FUNCTION_BLOCK TestingSequence (* Basic Function Block Type *)
  (* Standard: 61499-2 *)
  (* Version 0.0, 11/16/2026, Sandeep Patil, Flexbridge AB, Template *)
  PACKAGE Flexbridge.FestoMPS400;
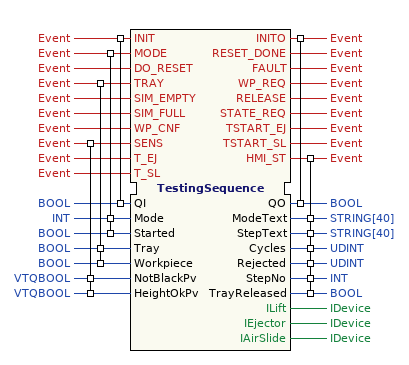
  EVENT_INPUT
    INIT WITH QI; (* Initialisation request *)
    MODE WITH Mode, Started; (* Station mode changed (StationMode) *)
    DO_RESET; (* Run the reset sequence (StationMode) *)
    TRAY WITH Tray, Workpiece; (* Tray state at interface 1 (conveyor waypoint, IWaypoint) *)
    SIM_EMPTY; (* Stand-in: an empty tray has arrived (HMI button) *)
    SIM_FULL; (* Stand-in: a tray with a workpiece has arrived (HMI button) *)
    WP_CNF; (* Distributing has handed a workpiece over (IWorkpieceSupply) *)
    SENS WITH NotBlackPv, HeightOkPv; (* Colour or height sensor changed *)
    T_EJ; (* Ejector time over (EjectTimer) *)
    T_SL; (* Air slide time over (SlideTimer) *)
  END_EVENT
  EVENT_OUTPUT
    INITO WITH QO; (* Initialisation confirm *)
    RESET_DONE; (* Reset sequence finished (StationMode) *)
    FAULT; (* Stopped on a device fault (StationMode) *)
    WP_REQ; (* Ask Distributing for a workpiece (IWorkpieceSupply) *)
    RELEASE; (* Release the tray (IWaypoint) *)
    STATE_REQ; (* Ask the waypoint for the tray state (IWaypoint) *)
    TSTART_EJ; (* Start the ejector timer *)
    TSTART_SL; (* Start the air slide timer *)
    HMI_ST WITH ModeText, StepText, Cycles, Rejected, StepNo, TrayReleased; (* State for the HMI *)
  END_EVENT
  VAR_INPUT
    QI : BOOL; (* Input event qualifier *)
    Mode : INT; (* Station mode: 0 = wait for RESET, 1 = resetting, 2 = wait for START, 3 = started *)
    Started : BOOL; (* Station started: trays are accepted *)
    Tray : BOOL; (* A tray is at the stopper of interface 1 *)
    Workpiece : BOOL; (* The tray carries a workpiece *)
    NotBlackPv : VTQBOOL; (* B2 workpiece is not black *)
    HeightOkPv : VTQBOOL; (* Height comparator: height correct *)
  END_VAR
  VAR_OUTPUT
    QO : BOOL; (* Output event qualifier *)
    ModeText : STRING[40]; (* Station mode as text *)
    StepText : STRING[40]; (* Current step as text (number and name) *)
    Cycles : UDINT; (* Workpieces put on a tray since start-up *)
    Rejected : UDINT; (* Workpieces rejected (black or wrong height) since start-up *)
    StepNo : INT; (* Current step number *)
    TrayReleased : BOOL; (* The tray has been released (until the next tray) *)
  END_VAR
  PLUGS
    ILift : IDevice;
    IEjector : IDevice;
    IAirSlide : IDevice;
  END_PLUGS
  VAR
    Done : BOOL; (* The current step has reached its target *)
    Fault : BOOL; (* A device needs Rearm, or is not program local when it must be *)
    Accept : BOOL; (* A tray is accepted (station started, tray present) *)
    TrayNow : BOOL; (* A tray is present (from the waypoint or a stand-in button) *)
    Full : BOOL; (* The present tray carries a workpiece *)
    Black : BOOL; (* The workpiece is black *)
    HeightGood : BOOL; (* The workpiece has the right height *)
    RdyLift : BOOL; (* Lift has sent CNF_READY: its owner has initialised *)
    AdpLift : BOOL; (* Lift taken over at start-up, or the reset sequence has run *)
    TryLift : INT; (* Program-local requests sent to Lift at start-up *)
  END_VAR
  EC_STATES
    START; (* Initial state *)
    INIT_S : algInit, algModeText, -> HMI_ST, -> INITO;
    S_IDLE : algModeText, algIdle -> HMI_ST;
    IDLE_W; (* Idle: wait for RESET (reset sequence) or a tray *)
    M_IDLE : algModeText -> HMI_ST;
    Q_TRAY : algQTray;
    Q_EMPTY : algQEmpty;
    Q_FULL : algQFull;
    Q_CHK : algQ_CHK;
    Q_NOSTART : algModeText -> HMI_ST;
    S_R_SEL : algModeText, algS_R_SEL -> HMI_ST, -> ILift.REQ_PROGLOCALSEL, -> IEjector.REQ_PROGLOCALSEL, -> IAirSlide.REQ_PROGLOCALSEL;
    C_R_SEL : algC_R_SEL;
    W_R_SEL; (* Wait: Reset: owners to program *)
    S_R_HOME : algModeText, algS_R_HOME -> HMI_ST, -> IAirSlide.REQ_CMD, -> ILift.REQ_CMD;
    C_R_HOME : algC_R_HOME;
    W_R_HOME; (* Wait: Reset: air off, lift down *)
    S_R_EJ : algModeText, algS_R_EJ -> HMI_ST, -> IEjector.REQ_CMD, -> TSTART_EJ;
    W_R_EJ; (* Wait: Reset: eject *)
    K_R_EJ : algFaultOnly;
    S_R_BACK : algModeText, algS_R_BACK -> HMI_ST, -> IEjector.REQ_CMD;
    C_R_BACK : algC_R_BACK;
    W_R_BACK; (* Wait: Reset: ejector back *)
    S_R_DONE : algModeText, algS_R_DONE -> HMI_ST, -> RESET_DONE, -> STATE_REQ;
    S_C_PASS : algModeText, algS_C_PASS -> HMI_ST, -> RELEASE;
    S_C_REQ : algModeText, algS_C_REQ -> HMI_ST, -> WP_REQ;
    W_C_REQ; (* Wait: Ask Distributing *)
    K_C_REQ : algFaultOnly;
    S_C_COLOUR : algModeText, algS_C_COLOUR -> HMI_ST;
    S_C_RAISE : algModeText, algS_C_RAISE -> HMI_ST, -> ILift.REQ_CMD;
    C_C_RAISE : algC_C_RAISE;
    W_C_RAISE; (* Wait: Raise lift *)
    S_C_HEIGHT : algModeText, algS_C_HEIGHT -> HMI_ST;
    S_C_PUSH : algModeText, algS_C_PUSH -> HMI_ST, -> IEjector.REQ_CMD, -> IAirSlide.REQ_CMD, -> TSTART_EJ;
    W_C_PUSH; (* Wait: Push onto air slide *)
    K_C_PUSH : algFaultOnly;
    S_C_BACK : algModeText, algS_C_BACK -> HMI_ST, -> IEjector.REQ_CMD;
    C_C_BACK : algC_C_BACK;
    W_C_BACK; (* Wait: Ejector back *)
    S_C_SLIDE : algModeText, algS_C_SLIDE -> HMI_ST, -> TSTART_SL;
    W_C_SLIDE; (* Wait: Air slide on *)
    K_C_SLIDE : algFaultOnly;
    S_C_LOWER : algModeText, algS_C_LOWER -> HMI_ST, -> IAirSlide.REQ_CMD, -> ILift.REQ_CMD;
    C_C_LOWER : algC_C_LOWER;
    W_C_LOWER; (* Wait: Air off, lift down *)
    S_C_DONE : algModeText, algS_C_DONE -> HMI_ST, -> RELEASE;
    S_X_LOWER : algModeText, algS_X_LOWER -> HMI_ST, -> ILift.REQ_CMD;
    C_X_LOWER : algC_X_LOWER;
    W_X_LOWER; (* Wait: Reject: lift down *)
    S_X_EJ : algModeText, algS_X_EJ -> HMI_ST, -> IEjector.REQ_CMD, -> TSTART_EJ;
    W_X_EJ; (* Wait: Reject: eject *)
    K_X_EJ : algFaultOnly;
    S_X_BACK : algModeText, algS_X_BACK -> HMI_ST, -> IEjector.REQ_CMD;
    C_X_BACK : algC_X_BACK;
    W_X_BACK; (* Wait: Reject: ejector back *)
    S_X_COUNT : algModeText, algS_X_COUNT -> HMI_ST;
    FAULT_S : algModeText, algFault -> HMI_ST, -> FAULT; (* Fault: RESET restarts the reset sequence after Rearm on the faceplate *)
    SR_Lift : algRdyLift; (* Lift ready before INIT *)
    TR_Lift : algRdyLift;
    TK_Lift; (* Start-up takeover of Lift *)
    TS_Lift : algTkSelLift -> ILift.REQ_PROGLOCALSEL;
    TC_Lift : algTkCmdLift -> ILift.REQ_CMD;
  END_STATES
  EC_TRANSITIONS
    START TO INIT_S := INIT;
    INIT_S TO S_IDLE := 1;
    S_IDLE TO TK_Lift := 1;
    IDLE_W TO INIT_S := INIT;
    IDLE_W TO M_IDLE := MODE;
    M_IDLE TO IDLE_W := 1;
    IDLE_W TO S_R_SEL := DO_RESET;
    IDLE_W TO Q_TRAY := TRAY;
    IDLE_W TO Q_EMPTY := SIM_EMPTY;
    IDLE_W TO Q_FULL := SIM_FULL;
    Q_TRAY TO Q_CHK := 1;
    Q_EMPTY TO Q_CHK := 1;
    Q_FULL TO Q_CHK := 1;
    Q_CHK TO Q_NOSTART := NOT Accept;
    Q_NOSTART TO IDLE_W := 1;
    Q_CHK TO FAULT_S := Accept AND Fault;
    Q_CHK TO S_C_PASS := Accept AND NOT Fault AND Full;
    Q_CHK TO S_C_REQ := Accept AND NOT Fault AND NOT Full;
    S_R_SEL TO C_R_SEL := 1;
    C_R_SEL TO FAULT_S := Fault;
    C_R_SEL TO S_R_HOME := NOT Fault AND Done;
    C_R_SEL TO W_R_SEL := NOT Fault AND NOT Done;
    W_R_SEL TO C_R_SEL := ILift.CNF_STATUS OR ILift.CNF_READY OR IEjector.CNF_STATUS OR IEjector.CNF_READY OR IAirSlide.CNF_STATUS OR IAirSlide.CNF_READY;
    S_R_HOME TO C_R_HOME := 1;
    C_R_HOME TO FAULT_S := Fault;
    C_R_HOME TO S_R_EJ := NOT Fault AND Done;
    C_R_HOME TO W_R_HOME := NOT Fault AND NOT Done;
    W_R_HOME TO C_R_HOME := ILift.CNF_STATUS OR ILift.CNF_READY OR IEjector.CNF_STATUS OR IEjector.CNF_READY OR IAirSlide.CNF_STATUS OR IAirSlide.CNF_READY;
    S_R_EJ TO W_R_EJ := 1;
    W_R_EJ TO S_R_BACK := T_EJ;
    W_R_EJ TO K_R_EJ := ILift.CNF_STATUS OR ILift.CNF_READY OR IEjector.CNF_STATUS OR IEjector.CNF_READY OR IAirSlide.CNF_STATUS OR IAirSlide.CNF_READY;
    K_R_EJ TO FAULT_S := Fault;
    K_R_EJ TO W_R_EJ := NOT Fault;
    S_R_BACK TO C_R_BACK := 1;
    C_R_BACK TO FAULT_S := Fault;
    C_R_BACK TO S_R_DONE := NOT Fault AND Done;
    C_R_BACK TO W_R_BACK := NOT Fault AND NOT Done;
    W_R_BACK TO C_R_BACK := ILift.CNF_STATUS OR ILift.CNF_READY OR IEjector.CNF_STATUS OR IEjector.CNF_READY OR IAirSlide.CNF_STATUS OR IAirSlide.CNF_READY;
    S_R_DONE TO IDLE_W := 1;
    S_C_PASS TO IDLE_W := 1;
    S_C_REQ TO W_C_REQ := 1;
    W_C_REQ TO S_C_COLOUR := WP_CNF;
    W_C_REQ TO K_C_REQ := ILift.CNF_STATUS OR ILift.CNF_READY OR IEjector.CNF_STATUS OR IEjector.CNF_READY OR IAirSlide.CNF_STATUS OR IAirSlide.CNF_READY;
    K_C_REQ TO FAULT_S := Fault;
    K_C_REQ TO W_C_REQ := NOT Fault;
    S_C_COLOUR TO S_X_EJ := Black;
    S_C_COLOUR TO S_C_RAISE := NOT Black;
    S_C_RAISE TO C_C_RAISE := 1;
    C_C_RAISE TO FAULT_S := Fault;
    C_C_RAISE TO S_C_HEIGHT := NOT Fault AND Done;
    C_C_RAISE TO W_C_RAISE := NOT Fault AND NOT Done;
    W_C_RAISE TO C_C_RAISE := ILift.CNF_STATUS OR ILift.CNF_READY OR IEjector.CNF_STATUS OR IEjector.CNF_READY OR IAirSlide.CNF_STATUS OR IAirSlide.CNF_READY;
    S_C_HEIGHT TO S_C_PUSH := HeightGood;
    S_C_HEIGHT TO S_X_LOWER := NOT HeightGood;
    S_C_PUSH TO W_C_PUSH := 1;
    W_C_PUSH TO S_C_BACK := T_EJ;
    W_C_PUSH TO K_C_PUSH := ILift.CNF_STATUS OR ILift.CNF_READY OR IEjector.CNF_STATUS OR IEjector.CNF_READY OR IAirSlide.CNF_STATUS OR IAirSlide.CNF_READY;
    K_C_PUSH TO FAULT_S := Fault;
    K_C_PUSH TO W_C_PUSH := NOT Fault;
    S_C_BACK TO C_C_BACK := 1;
    C_C_BACK TO FAULT_S := Fault;
    C_C_BACK TO S_C_SLIDE := NOT Fault AND Done;
    C_C_BACK TO W_C_BACK := NOT Fault AND NOT Done;
    W_C_BACK TO C_C_BACK := ILift.CNF_STATUS OR ILift.CNF_READY OR IEjector.CNF_STATUS OR IEjector.CNF_READY OR IAirSlide.CNF_STATUS OR IAirSlide.CNF_READY;
    S_C_SLIDE TO W_C_SLIDE := 1;
    W_C_SLIDE TO S_C_LOWER := T_SL;
    W_C_SLIDE TO K_C_SLIDE := ILift.CNF_STATUS OR ILift.CNF_READY OR IEjector.CNF_STATUS OR IEjector.CNF_READY OR IAirSlide.CNF_STATUS OR IAirSlide.CNF_READY;
    K_C_SLIDE TO FAULT_S := Fault;
    K_C_SLIDE TO W_C_SLIDE := NOT Fault;
    S_C_LOWER TO C_C_LOWER := 1;
    C_C_LOWER TO FAULT_S := Fault;
    C_C_LOWER TO S_C_DONE := NOT Fault AND Done;
    C_C_LOWER TO W_C_LOWER := NOT Fault AND NOT Done;
    W_C_LOWER TO C_C_LOWER := ILift.CNF_STATUS OR ILift.CNF_READY OR IEjector.CNF_STATUS OR IEjector.CNF_READY OR IAirSlide.CNF_STATUS OR IAirSlide.CNF_READY;
    S_C_DONE TO IDLE_W := 1;
    S_X_LOWER TO C_X_LOWER := 1;
    C_X_LOWER TO FAULT_S := Fault;
    C_X_LOWER TO S_X_EJ := NOT Fault AND Done;
    C_X_LOWER TO W_X_LOWER := NOT Fault AND NOT Done;
    W_X_LOWER TO C_X_LOWER := ILift.CNF_STATUS OR ILift.CNF_READY OR IEjector.CNF_STATUS OR IEjector.CNF_READY OR IAirSlide.CNF_STATUS OR IAirSlide.CNF_READY;
    S_X_EJ TO W_X_EJ := 1;
    W_X_EJ TO S_X_BACK := T_EJ;
    W_X_EJ TO K_X_EJ := ILift.CNF_STATUS OR ILift.CNF_READY OR IEjector.CNF_STATUS OR IEjector.CNF_READY OR IAirSlide.CNF_STATUS OR IAirSlide.CNF_READY;
    K_X_EJ TO FAULT_S := Fault;
    K_X_EJ TO W_X_EJ := NOT Fault;
    S_X_BACK TO C_X_BACK := 1;
    C_X_BACK TO FAULT_S := Fault;
    C_X_BACK TO S_X_COUNT := NOT Fault AND Done;
    C_X_BACK TO W_X_BACK := NOT Fault AND NOT Done;
    W_X_BACK TO C_X_BACK := ILift.CNF_STATUS OR ILift.CNF_READY OR IEjector.CNF_STATUS OR IEjector.CNF_READY OR IAirSlide.CNF_STATUS OR IAirSlide.CNF_READY;
    S_X_COUNT TO S_C_REQ := 1;
    FAULT_S TO IDLE_W := 1;
    START TO SR_Lift := ILift.CNF_READY;
    SR_Lift TO START := 1;
    IDLE_W TO TR_Lift := ILift.CNF_READY;
    TR_Lift TO TK_Lift := 1;
    IDLE_W TO TK_Lift := ILift.CNF_STATUS;
    TK_Lift TO TS_Lift := NOT AdpLift AND RdyLift AND NOT ILift.ProgLocal AND TryLift < 3;
    TK_Lift TO TC_Lift := NOT AdpLift AND RdyLift AND ILift.ProgLocal AND (ILift.Status.value = 1 OR ILift.Status.value = 2);
    TK_Lift TO IDLE_W := NOT (NOT AdpLift AND RdyLift AND NOT ILift.ProgLocal AND TryLift < 3) AND NOT (NOT AdpLift AND RdyLift AND ILift.ProgLocal AND (ILift.Status.value = 1 OR ILift.Status.value = 2));
    TS_Lift TO IDLE_W := 1;
    TC_Lift TO IDLE_W := 1;
  END_TRANSITIONS
  ALGORITHM algModeText IN ST: (* Station mode as text *)
CASE Mode OF
    0: ModeText := 'Wait for RESET';
    1: ModeText := 'Resetting';
    2: ModeText := 'Wait for START';
    3: ModeText := 'Started';
ELSE
    ModeText := 'Unknown mode';
END_CASE;
  END_ALGORITHM
  ALGORITHM algInit IN ST: (* Idle *)
QO := QI;
StepNo := 0; StepText := '0 Idle';
Cycles := 0; Rejected := 0; TrayReleased := FALSE;
Done := FALSE; Fault := FALSE;
AdpLift := FALSE; TryLift := 0;
  END_ALGORITHM
  ALGORITHM algIdle IN ST: (* Idle *)
StepNo := 0; StepText := '0 Idle';
  END_ALGORITHM
  ALGORITHM algFaultOnly IN ST: (* Fault check while waiting for a timer or a confirmation *)
Fault := ILift.NeedReset OR IEjector.NeedReset OR IAirSlide.NeedReset;
  END_ALGORITHM
  ALGORITHM algQTray IN ST: (* Tray state from the waypoint *)
TrayNow := Tray; Full := Workpiece;
  END_ALGORITHM
  ALGORITHM algQEmpty IN ST: (* Stand-in: empty tray *)
TrayNow := TRUE; Full := FALSE;
  END_ALGORITHM
  ALGORITHM algQFull IN ST: (* Stand-in: tray with a workpiece *)
TrayNow := TRUE; Full := TRUE;
  END_ALGORITHM
  ALGORITHM algQ_CHK IN ST: (* Tray: accept only when started; all devices must be ready *)
Accept := Started AND TrayNow;
Fault := ILift.NeedReset OR IEjector.NeedReset OR IAirSlide.NeedReset OR NOT (ILift.ProgLocal AND IEjector.ProgLocal AND IAirSlide.ProgLocal);
IF NOT Started THEN
    StepText := '0 Idle: press START first';
ELSIF NOT TrayNow THEN
    StepText := '0 Idle: no tray';
END_IF;
  END_ALGORITHM
  ALGORITHM algS_R_SEL IN ST: (* Reset: owners to program *)
StepNo := 10; StepText := '10 Reset: owners to program';
ILift.ProgLocalSel := TRUE;
IEjector.ProgLocalSel := TRUE;
IAirSlide.ProgLocalSel := TRUE;
AdpLift := TRUE;
  END_ALGORITHM
  ALGORITHM algC_R_SEL IN ST: (* Check: Reset: owners to program *)
Fault := ILift.NeedReset OR IEjector.NeedReset OR IAirSlide.NeedReset;
Done := ILift.ProgLocal AND IEjector.ProgLocal AND IAirSlide.ProgLocal;
  END_ALGORITHM
  ALGORITHM algS_R_HOME IN ST: (* Reset: air off, lift down *)
StepNo := 11; StepText := '11 Reset: air off, lift down';
IAirSlide.Lsp.value := 0;
ILift.Lsp.value := 2;
  END_ALGORITHM
  ALGORITHM algC_R_HOME IN ST: (* Check: Reset: air off, lift down *)
Fault := ILift.NeedReset OR IEjector.NeedReset OR IAirSlide.NeedReset;
Done := ILift.Status.value = 2;
  END_ALGORITHM
  ALGORITHM algS_R_EJ IN ST: (* Reset: eject *)
StepNo := 12; StepText := '12 Reset: eject';
IEjector.Lsp.value := 1;
  END_ALGORITHM
  ALGORITHM algS_R_BACK IN ST: (* Reset: ejector back *)
StepNo := 13; StepText := '13 Reset: ejector back';
IEjector.Lsp.value := 2;
  END_ALGORITHM
  ALGORITHM algC_R_BACK IN ST: (* Check: Reset: ejector back *)
Fault := ILift.NeedReset OR IEjector.NeedReset OR IAirSlide.NeedReset;
Done := IEjector.Status.value = 2;
  END_ALGORITHM
  ALGORITHM algS_R_DONE IN ST: (* Reset done *)
StepNo := 14; StepText := '14 Reset done';
TrayReleased := FALSE;
  END_ALGORITHM
  ALGORITHM algS_C_PASS IN ST: (* Tray full: released *)
StepNo := 20; StepText := '20 Tray full: released';
TrayReleased := TRUE;
  END_ALGORITHM
  ALGORITHM algS_C_REQ IN ST: (* Ask Distributing *)
StepNo := 21; StepText := '21 Ask Distributing';
TrayReleased := FALSE;
  END_ALGORITHM
  ALGORITHM algS_C_COLOUR IN ST: (* Check colour *)
StepNo := 22; StepText := '22 Check colour';
Black := NOT NotBlackPv.value;
  END_ALGORITHM
  ALGORITHM algS_C_RAISE IN ST: (* Raise lift *)
StepNo := 23; StepText := '23 Raise lift';
ILift.Lsp.value := 1;
  END_ALGORITHM
  ALGORITHM algC_C_RAISE IN ST: (* Check: Raise lift *)
Fault := ILift.NeedReset OR IEjector.NeedReset OR IAirSlide.NeedReset;
Done := ILift.Status.value = 1;
  END_ALGORITHM
  ALGORITHM algS_C_HEIGHT IN ST: (* Check height *)
StepNo := 24; StepText := '24 Check height';
HeightGood := HeightOkPv.value;
  END_ALGORITHM
  ALGORITHM algS_C_PUSH IN ST: (* Push onto air slide *)
StepNo := 25; StepText := '25 Push onto air slide';
IEjector.Lsp.value := 1;
IAirSlide.Lsp.value := 1;
  END_ALGORITHM
  ALGORITHM algS_C_BACK IN ST: (* Ejector back *)
StepNo := 26; StepText := '26 Ejector back';
IEjector.Lsp.value := 2;
  END_ALGORITHM
  ALGORITHM algC_C_BACK IN ST: (* Check: Ejector back *)
Fault := ILift.NeedReset OR IEjector.NeedReset OR IAirSlide.NeedReset;
Done := IEjector.Status.value = 2;
  END_ALGORITHM
  ALGORITHM algS_C_SLIDE IN ST: (* Air slide on *)
StepNo := 27; StepText := '27 Air slide on';
  END_ALGORITHM
  ALGORITHM algS_C_LOWER IN ST: (* Air off, lift down *)
StepNo := 28; StepText := '28 Air off, lift down';
IAirSlide.Lsp.value := 0;
ILift.Lsp.value := 2;
  END_ALGORITHM
  ALGORITHM algC_C_LOWER IN ST: (* Check: Air off, lift down *)
Fault := ILift.NeedReset OR IEjector.NeedReset OR IAirSlide.NeedReset;
Done := ILift.Status.value = 2;
  END_ALGORITHM
  ALGORITHM algS_C_DONE IN ST: (* Done: tray released *)
StepNo := 29; StepText := '29 Done: tray released';
Cycles := Cycles + 1;
TrayReleased := TRUE;
  END_ALGORITHM
  ALGORITHM algS_X_LOWER IN ST: (* Reject: lift down *)
StepNo := 32; StepText := '32 Reject: lift down';
ILift.Lsp.value := 2;
  END_ALGORITHM
  ALGORITHM algC_X_LOWER IN ST: (* Check: Reject: lift down *)
Fault := ILift.NeedReset OR IEjector.NeedReset OR IAirSlide.NeedReset;
Done := ILift.Status.value = 2;
  END_ALGORITHM
  ALGORITHM algS_X_EJ IN ST: (* Reject: eject *)
StepNo := 30; StepText := '30 Reject: eject';
IEjector.Lsp.value := 1;
  END_ALGORITHM
  ALGORITHM algS_X_BACK IN ST: (* Reject: ejector back *)
StepNo := 31; StepText := '31 Reject: ejector back';
IEjector.Lsp.value := 2;
  END_ALGORITHM
  ALGORITHM algC_X_BACK IN ST: (* Check: Reject: ejector back *)
Fault := ILift.NeedReset OR IEjector.NeedReset OR IAirSlide.NeedReset;
Done := IEjector.Status.value = 2;
  END_ALGORITHM
  ALGORITHM algS_X_COUNT IN ST: (* Rejected: ask again *)
StepNo := 33; StepText := '33 Rejected: ask again';
Rejected := Rejected + 1;
  END_ALGORITHM
  ALGORITHM algFault IN ST: (* Device fault: stop here, report to StationMode *)
StepNo := 99;
IF ILift.NeedReset THEN
    StepText := '99 FAULT: Rearm Lift';
ELSIF IEjector.NeedReset THEN
    StepText := '99 FAULT: Rearm Ejector';
ELSIF IAirSlide.NeedReset THEN
    StepText := '99 FAULT: Rearm AirSlide';
ELSE
    StepText := '99 FAULT: owner not program';
END_IF;
  END_ALGORITHM
  ALGORITHM algRdyLift IN ST: (* Lift has reported ready *)
RdyLift := TRUE;
  END_ALGORITHM
  ALGORITHM algTkSelLift IN ST: (* Start-up: ask Lift for program local *)
ILift.ProgLocalSel := TRUE;
TryLift := TryLift + 1;
  END_ALGORITHM
  ALGORITHM algTkCmdLift IN ST: (* Start-up: command the end position Lift reports (it does not move) *)
ILift.Lsp.value := ILift.Status.value;
AdpLift := TRUE;
  END_ALGORITHM
END_FUNCTION_BLOCK
